// TIA Portal V21 export
FUNCTION_BLOCK "Mixed"   // FB12, LAD
TITLE = Mixed languages
{ S7_Optimized_Access := 'TRUE' }
// A ladder block with an SCL and an STL network.
   VAR_INPUT
      start : Bool;
      stop : Bool;
      door : Bool;
   END_VAR
   VAR_OUTPUT
      motor : Bool;
      lamp : Bool;
      fault : Bool;
   END_VAR
   VAR
      latched : Bool;
      edgeMemory : Bool;
   END_VAR
BEGIN

REGION Network 1: Ladder
   // A ladder network first.
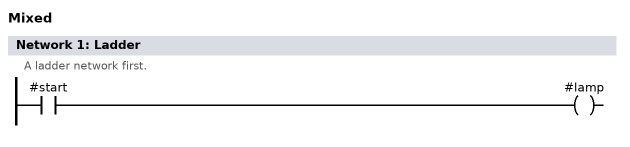
   RUNG wire#powerrail
      Contact( #start )
      Coil( #lamp )
   END_RUNG
   // the same network as SCL:
   #lamp := #start;
END_REGION

REGION Network 2 (SCL): Structured text
   // An SCL network inside a ladder block.
   #motor := #start AND NOT #stop;
END_REGION

NETWORK
TITLE = Statement list
// An STL network inside a ladder block.
      A     #door;
      AN    #stop;
      =     #fault;
END_FUNCTION_BLOCK
